(* IEC 61131-3 sources: axsharp/src/sanbox/probes/ax-blazor-1/src, 4 files *)

(* ---- geolocation.st ---- *)
{ix:[Container(Layout.Stack)]}
{ix:[Group(Layout.GroupBox, "GEOLOCATION")]}
CLASS  GeoLocation
    VAR PUBLIC
        Latitude : REAL;
        Longitude : REAL;
        Altitude : REAL;
        Description : STRING;
    END_VAR
END_CLASS

(* ---- weather.st ---- *)
CLASS weather
    VAR PUBLIC
        Temperature : REAL;
        Humidity : REAL;
        Location : STRING;
        HeyMan : STRING;
        GeoLocation : GeoLocation;
    END_VAR
END_CLASS

CLASS weathers
    VAR PUBLIC
        i : ARRAY[0..10] OF weather;
    END_VAR
END_CLASS

(* ---- configuration.st ---- *)
CONFIGURATION MyConfiguration
    TASK Main(Interval := T#1000ms, Priority := 1);
    PROGRAM P1 WITH Main: MyProgram;

    VAR_GLOBAL
        myINT : INT;
        weather : weather;
        weathers : weathers;
    END_VAR
END_CONFIGURATION

(* ---- program.st ---- *)
PROGRAM MyProgram
    VAR_EXTERNAL
        myINT : INT;
    END_VAR

    VAR

    END_VAR

    VAR_TEMP

    END_VAR

    myINT := myINT + 1;
END_PROGRAM
